// TIA Portal V21 export
// export: Created 2026-08-21T20:18:50.9872746Z, ExportSetting None, DisplayName Totally Integrated Automation Portal, DisplayVersion V21, DisplayName STEP 7 Professional, DisplayVersion V21, DisplayName STEP 7 Safety, DisplayVersion V21, DisplayName Tech WebApplication, DisplayVersion V21, DisplayName WinCC Basic/Comfort/Advanced, DisplayVersion V21, DisplayName WinCC Professional, DisplayVersion V21, DisplayName WinCC Unified, DisplayVersion V21
FUNCTION "P100" : Void   // FC2, FBD
{ S7_Optimized_Access := 'TRUE' }
// stored: SetENOAutomatically false
   VAR_TEMP
      Temp : "DigVal";
      Temp_1 : "DigVal";
      Temp_3 : "DigVal";
      Temp_2 : "DigVal";
      Temp_Error : "DigVal";
      In03 : "DigVal";
      State : "Service_States";
      FbkRun : "DigVal";
      StopAut : Bool;
   END_VAR
   VAR_TEMP   // added for the SCL form of the ladder/FBD networks
      _w1 : Bool;
   END_VAR
BEGIN

REGION Network 1: simulate Fbk Error
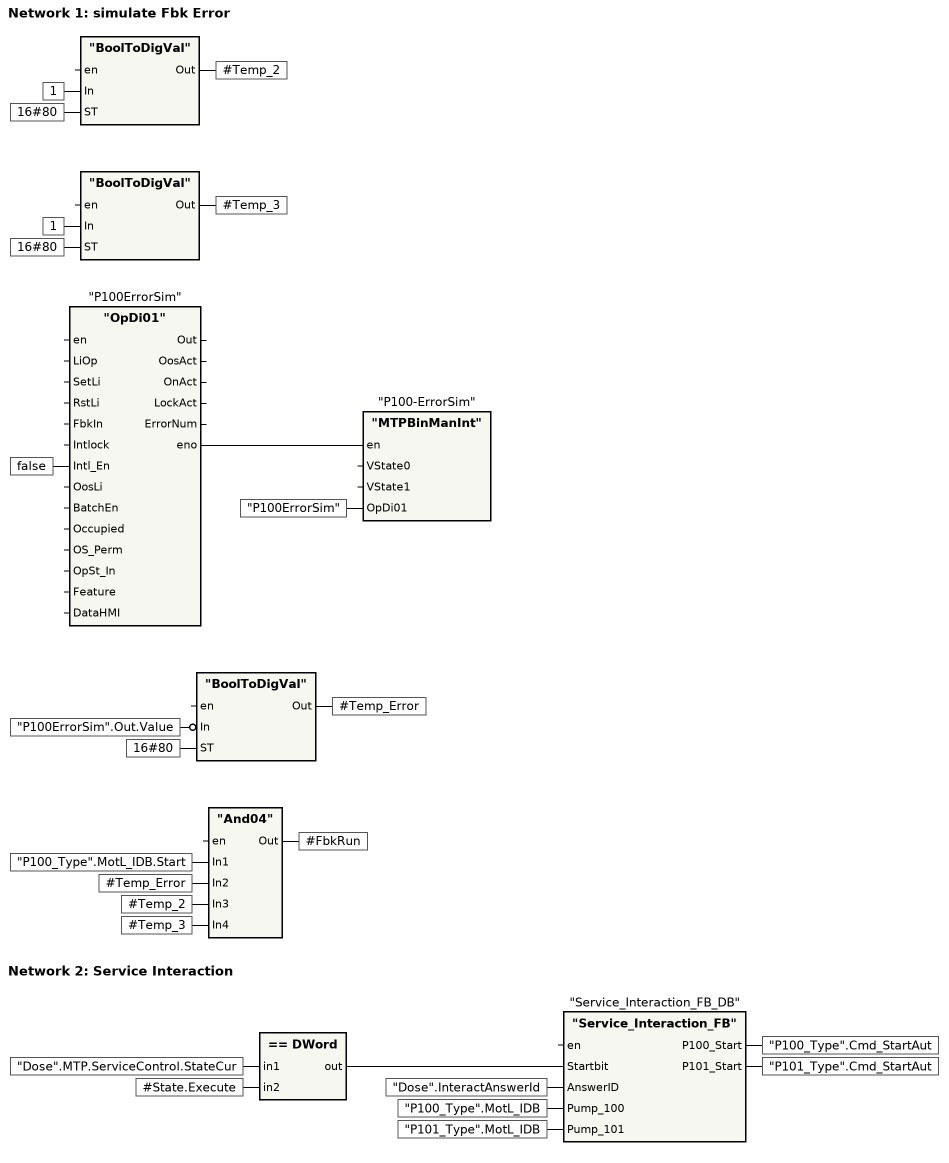
   "BoolToDigVal"(In := 1, ST := 16#80, Out => #Temp_2);
   "BoolToDigVal"(In := 1, ST := 16#80, Out => #Temp_3);
   "P100ErrorSim"(Intl_En := false, ENO => #_w1);   // "OpDi01"
   IF #_w1 THEN
       "P100-ErrorSim"(OpDi01 := "P100ErrorSim");   // "MTPBinManInt"
   END_IF;
   "BoolToDigVal"(In := NOT "P100ErrorSim".Out.Value, ST := 16#80, Out => #Temp_Error);
   "And04"(In1 := "P100_Type".MotL_IDB.Start,
           In2 := #Temp_Error,
           In3 := #Temp_2,
           In4 := #Temp_3,
           Out => #FbkRun);
END_REGION

REGION Network 2: Service Interaction
   "Service_Interaction_FB_DB"(Startbit := "Dose".MTP.ServiceControl.StateCur = #State.Execute,   // "Service_Interaction_FB"
                           AnswerID := "Dose".InteractAnswerId,
                           Pump_100 := "P100_Type".MotL_IDB,
                           Pump_101 := "P101_Type".MotL_IDB,
                           P100_Start => "P100_Type".Cmd_StartAut,
                           P101_Start => "P101_Type".Cmd_StartAut);
END_REGION

REGION Network 3: Pump interconnections
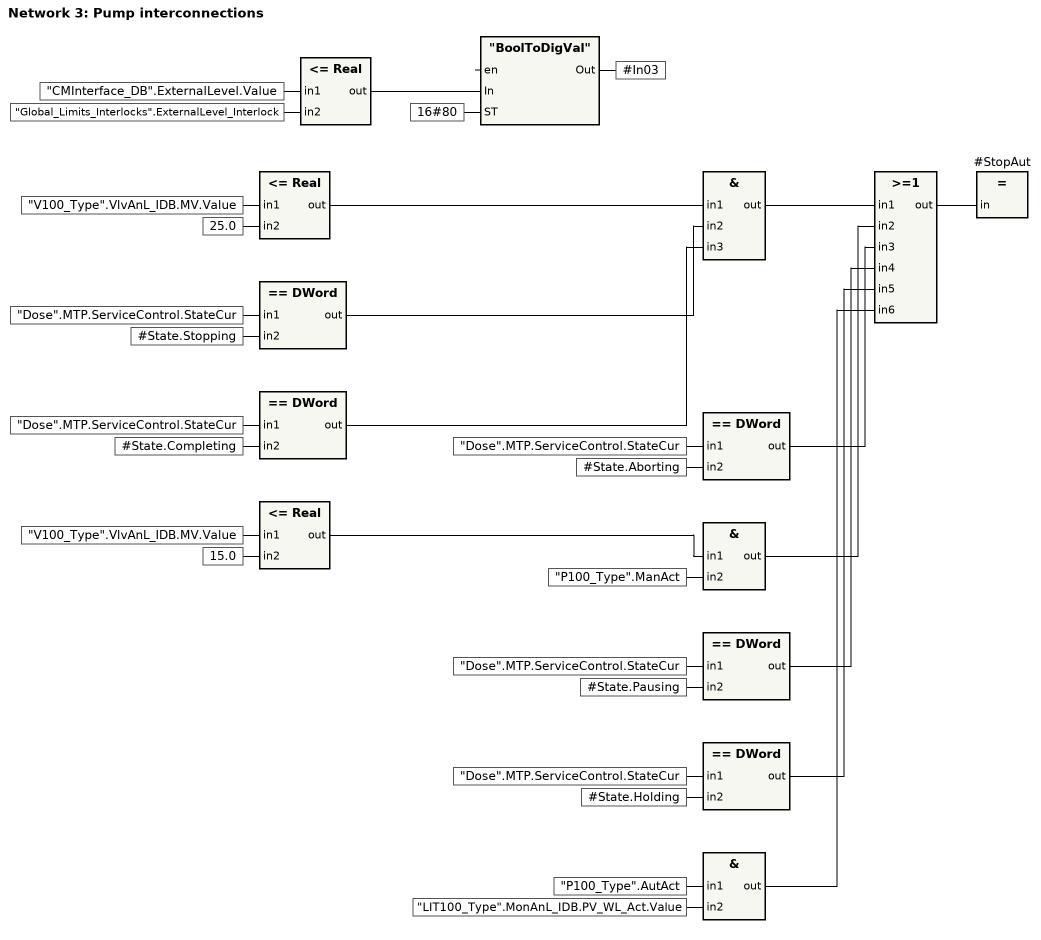
   "BoolToDigVal"(In := "CMInterface_DB".ExternalLevel.Value <= "Global_Limits_Interlocks".ExternalLevel_Interlock,
                  ST := 16#80,
                  Out => #In03);
   #StopAut := (("V100_Type".VlvAnL_IDB.MV.Value <= 25.0) AND ("Dose".MTP.ServiceControl.StateCur = #State.Stopping) AND ("Dose".MTP.ServiceControl.StateCur = #State.Completing)) OR (("V100_Type".VlvAnL_IDB.MV.Value <= 15.0) AND "P100_Type".ManAct) OR ("Dose".MTP.ServiceControl.StateCur = #State.Aborting) OR ("Dose".MTP.ServiceControl.StateCur = #State.Pausing) OR ("Dose".MTP.ServiceControl.StateCur = #State.Holding) OR ("P100_Type".AutAct AND "LIT100_Type".MonAnL_IDB.PV_WL_Act.Value);
END_REGION

REGION Network 4: MotL
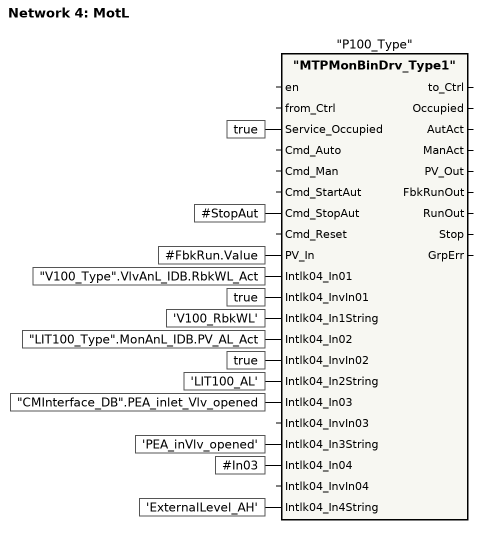
   "P100_Type"(Service_Occupied := true,   // "MTPMonBinDrv_Type1"
               Cmd_StopAut := #StopAut,
               PV_In := #FbkRun.Value,
               Intlk04_In01 := "V100_Type".VlvAnL_IDB.RbkWL_Act,
               Intlk04_InvIn01 := true,
               Intlk04_In1String := 'V100_RbkWL',
               Intlk04_In02 := "LIT100_Type".MonAnL_IDB.PV_AL_Act,
               Intlk04_InvIn02 := true,
               Intlk04_In2String := 'LIT100_AL',
               Intlk04_In03 := "CMInterface_DB".PEA_inlet_Vlv_opened,
               Intlk04_In3String := 'PEA_inVlv_opened',
               Intlk04_In04 := #In03,
               Intlk04_In4String := 'ExternalLevel_AH');
END_REGION
END_FUNCTION
